{region 'Documentation'}
(*!
<summary>Checks an individually impossible execution budget against actual usable capacity.</summary>
<description>

Real subject boundaries

The real Test Case computes reservations; the real Orchestrator decides and publishes its diagnostic.
A collection double supplies one fixed child view. Only the concurrent Suite allowance is held by
the fixture, without running a Suite. Request-entry observations are inherited from the thin child adapter.
The physical array includes one unused FIFO position, leaving capacity one entry below the minimum.
The buffer is empty at rejection: consumer deletion cannot repair an impossible budget.
Three later helper calls must retain Error without another diagnostic or unexpected dispatch.
Expected diagnostics stay in local capture. The surrounding Assertions use the normal selftest publisher.
The real subject binds only local storage; expected findings remain in that storage.
Checking Assertions retain the outer selftest publisher. Each run reinitializes the subject.
</description>
*)
{endregion}
FUNCTION_BLOCK Test_ImpossibleExecutionBudget EXTENDS TestCaseBase
VAR
    FSubject : EventBuffer;
    FEvents : ARRAY[1..BufferLength] OF ST_Event;
    FFifo : ST_FifoStatus;
    FBufferStatus : ST_EventBufferStatus;
    FPerformed : BOOL;
    FChecked : BOOL;
    FSubjectParent : I_TestSuite;
    FChild : ReservationChildProbe;
    FOrchestrator : OrchestratorProbe;
    FCollection : OrchestrationCollectionDouble;
    FChildren : ARRAY[1..1] OF I_Orchestratable;
    FOwnerReserved : UINT;
    FStep : INT;
    FObservationCalls : UINT;
    FPrecondition : AssertTrue;
    FPreconditionMatches : BOOL;
    FFailureDetection : AssertTrue;
    FFailureDetectionMatches : BOOL;
    FStateAndCounts : AssertTrue;
    FStateAndCountsMatches : BOOL;
    FHeldError : AssertTrue;
    FHeldErrorMatches : BOOL;
    FSingleDiagnostic : AssertTrue;
    FSingleDiagnosticMatches : BOOL;
    FRequestBoundary : AssertTrue;
    FRequestBoundaryMatches : BOOL;
    FAccounting : AssertTrue;
    FAccountingMatches : BOOL;
    FCaptureIntegrity : AssertTrue;
    FCaptureIntegrityMatches : BOOL;
END_VAR
VAR CONSTANT
    ChildExecutionBudget : UINT := 11;
    ConfigureExecution : INT := 4;
    BufferLength : UINT := GVL_Constants.TestSuiteExecutionEventCount + ChildExecutionBudget + Param_EventBuffer.EventBufferExecutionHeadroom;
    ObservationCalls : UINT := 3;
    ExpectedResetRequests : UINT := 1;
    ExpectedStartRequests : UINT := 0;
    Setup : INT := 0;
    PrepareChild : INT := 1;
    TriggerFailure : INT := 2;
    ObserveFailure : INT := 3;
END_VAR

SUPER^();

{region 'Documentation'}
(*!
<summary>Contributes each checking Assertion once.</summary>
*)
{endregion}
METHOD PROTECTED AggregateResults
VAR_INPUT
    Aggregator : I_ResultAggregator; //! Borrowed result sink owned by the outer Test Case; add this test's checking Assertions without resetting or retaining the sink.
END_VAR
Aggregator.AddProvider(Provider := FPrecondition);
Aggregator.AddProvider(Provider := FFailureDetection);
Aggregator.AddProvider(Provider := FStateAndCounts);
Aggregator.AddProvider(Provider := FHeldError);
Aggregator.AddProvider(Provider := FSingleDiagnostic);
Aggregator.AddProvider(Provider := FRequestBoundary);
Aggregator.AddProvider(Provider := FAccounting);
Aggregator.AddProvider(Provider := FCaptureIntegrity);
END_METHOD

{region 'Documentation'}
(*!
<summary>Supplies only the child identity before initialization.</summary>
*)
{endregion}
METHOD PUBLIC BindSubjectParent
VAR_INPUT
    Parent : I_TestSuite; //! Borrowed identity parent retained for isolated subject initialization; keep the Suite alive through subject use.
END_VAR
FSubjectParent := Parent;
END_METHOD

{region 'Documentation'}
(*!
<summary>Calls the real helper and child and retains accounting observations.</summary>
*)
{endregion}
METHOD PRIVATE CallSubject
VAR_INPUT
    Task : E_OrchestratorTask; //! Orchestration task assigned for this controlled subject call.
END_VAR
FOrchestrator(Task := Task);
FAccountingMatches := FAccountingMatches
    AND (FSubject.ReservedEntryCount = FOwnerReserved + FChild.ReservedEntryCount);
FChild();
FCaptureIntegrityMatches := FCaptureIntegrityMatches
    AND NOT FFifo.ConfigError AND NOT FFifo.IndexError
    AND (FBufferStatus.LostEventCount = 0)
    AND NOT FCollection.InvalidAccess AND NOT FCollection.TraceOverflow;
END_METHOD

{region 'Documentation'}
(*!
<summary>Checks the single retained Orchestrator Error and exact dispatch counts.</summary>
*)
{endregion}
METHOD PRIVATE CheckDiagnostic
VAR
    Index : UINT;
    ErrorCount : UINT;
    PayloadMatches : BOOL := TRUE;
END_VAR
FOR Index := 1 TO BufferLength DO
    IF (FEvents[Index].SequenceId > 0) AND (FEvents[Index].Severity = E_EventSeverity.Error) THEN
        ErrorCount := ErrorCount + 1;
        PayloadMatches := PayloadMatches
            AND (FEvents[Index].OwnerScope = E_OwnerScope.Framework)
            AND (FEvents[Index].EventType = E_EventType.Framework)
            AND (FEvents[Index].State = E_State.Error)
            AND (FEvents[Index].Name = CONCAT(Name, '.Orchestrator'))
            AND (FEvents[Index].Message <> '');
    END_IF;
END_FOR;
FSingleDiagnosticMatches := (ErrorCount = 1) AND PayloadMatches;
FRequestBoundaryMatches := FChild.RequestsReserved
    AND (FChild.ResetRequestCount = ExpectedResetRequests)
    AND (FChild.StartRequestCount = ExpectedStartRequests);
END_METHOD

{region 'Documentation'}
(*!
<summary>Requires all checking Assertions to be initialized.</summary>
*)
{endregion}
METHOD PROTECTED CheckInitialization : BOOL //! TRUE when the inherited initialization check and this concrete fixture check both accept the setup.
CheckInitialization := FALSE;
IF NOT SUPER^.CheckInitialization() OR (FSubjectParent = 0) THEN
    RETURN;
END_IF;

CheckInitialization := FPrecondition.IsInitialized
    AND FFailureDetection.IsInitialized
    AND FStateAndCounts.IsInitialized
    AND FHeldError.IsInitialized
    AND FSingleDiagnostic.IsInitialized
    AND FRequestBoundary.IsInitialized
    AND FAccounting.IsInitialized
    AND FCaptureIntegrity.IsInitialized;
END_METHOD

{region 'Documentation'}
(*!
<summary>Initializes the checking Assertions for one test state.</summary>
*)
{endregion}
METHOD PROTECTED Configure
FPreparationStateCount := 0;
FTestStateCount := 1;
FPrecondition.Initialize(Parent := THIS^,
    AssertionName := 'Precondition');
FFailureDetection.Initialize(Parent := THIS^,
    AssertionName := 'FailureDetection');
FStateAndCounts.Initialize(Parent := THIS^,
    AssertionName := 'StateAndCounts');
FHeldError.Initialize(Parent := THIS^,
    AssertionName := 'HeldError');
FSingleDiagnostic.Initialize(Parent := THIS^,
    AssertionName := 'SingleDiagnostic');
FRequestBoundary.Initialize(Parent := THIS^,
    AssertionName := 'RequestBoundary');
FAccounting.Initialize(Parent := THIS^,
    AssertionName := 'Accounting');
FCaptureIntegrity.Initialize(Parent := THIS^,
    AssertionName := 'CaptureIntegrity');
END_METHOD

{region 'Documentation'}
(*!
<summary>Binds a real child and Orchestrator to fixed isolated storage.</summary>
*)
{endregion}
METHOD PRIVATE InitializeArrangement
VAR
    Config : ST_TestCaseConfig;
END_VAR
IF NOT FSubject.Initialize(Buffer := FEvents,
    FifoControl := FFifo,
    Status := FBufferStatus) THEN
    Error(Message := 'Reservation error capture initialization failed.');
    RETURN;
END_IF;
FOwnerReserved := 0;
FChild.BindPublisher(Publisher := FSubject);
FChild.ClearRequestTrace();
FChild.ExecutionSlot := 1;
IF NOT FChild.Initialize(Parent := FSubjectParent,
    TestName := 'ExecutionBudgetChild',
    Config := Config) THEN
    Error(Message := 'Reservation error child initialization failed.');
    RETURN;
END_IF;
FChild();
FChildren[1] := FChild;
IF NOT FCollection.Initialize(Count := 1,
    Children := FChildren) THEN
    Error(Message := 'Reservation error collection initialization failed.');
    RETURN;
END_IF;
FOrchestrator.BindPublisher(Publisher := FSubject);
IF NOT FOrchestrator.Initialize(Collection := FCollection,
    Name := Name) THEN
    Error(Message := 'Reservation error Orchestrator initialization failed.');
    RETURN;
END_IF;
IF NOT FSubject.ReserveSpace(EntryCount := GVL_Constants.TestSuiteResetEventCount,
    HeadroomEntryCount := Param_EventBuffer.EventBufferResetHeadroom,
    OwnerReservedEntryCount := FOwnerReserved) THEN
    Error(Message := 'Reservation error concurrent owner setup failed.');
    RETURN;
END_IF;
FPreconditionMatches := FPreconditionMatches AND FChild.IsInitialized
    AND FFifo.BufferEmpty AND (FSubject.Capacity = BufferLength - 1);
END_METHOD

{region 'Documentation'}
(*!
<summary>Removes setup events and replaces the fixture owner allowance; child configuration remains unchanged.</summary>
*)
{endregion}
METHOD PRIVATE PrepareExecution
VAR
    Watermark : UDINT;
END_VAR
Watermark := FBufferStatus.SequenceId;
FSubject.ProcessDeleteRequest(SequenceId := Watermark);
IF NOT FSubject.FreeReservedSpace(EntryCount := FOwnerReserved,
    OwnerReservedEntryCount := FOwnerReserved) THEN
    Error(Message := 'Could not release Reset fixture allowance.');
    RETURN;
END_IF;
IF NOT FSubject.ReserveSpace(EntryCount := GVL_Constants.TestSuiteExecutionEventCount,
    HeadroomEntryCount := Param_EventBuffer.EventBufferExecutionHeadroom,
    OwnerReservedEntryCount := FOwnerReserved) THEN
    Error(Message := 'Could not reserve execution fixture allowance.');
    RETURN;
END_IF;
FPreconditionMatches := FPreconditionMatches AND FFifo.BufferEmpty
    AND (Watermark = 0) AND (FChild.ReservedEntryCount = 0);
END_METHOD

{region 'Documentation'}
(*!
<summary>Completes abort without asynchronous work.</summary>
*)
{endregion}
METHOD PROTECTED ProcessAbort
VAR_INPUT
    Enable : BOOL; //! Phase permission supplied by the owning Test Case; FALSE does not authorize progression, while observation may continue.
END_VAR
IF Enable THEN
    CompleteAbort();
END_IF;
END_METHOD

{region 'Documentation'}
(*!
<summary>Evaluates captured observations after the scenario has finished.</summary>
*)
{endregion}
METHOD PROTECTED ProcessAssertions
VAR_INPUT
    Enable : BOOL; //! Phase permission supplied by the owning Test Case; FALSE does not authorize progression, while observation may continue.
END_VAR
VAR
    Evaluate : BOOL;
END_VAR
Evaluate := Enable AND FPerformed;
FPrecondition(Enable := Evaluate,
    State := State,
    IN := FPreconditionMatches);
FFailureDetection(Enable := Evaluate,
    State := State,
    IN := FFailureDetectionMatches);
FStateAndCounts(Enable := Evaluate,
    State := State,
    IN := FStateAndCountsMatches);
FHeldError(Enable := Evaluate,
    State := State,
    IN := FHeldErrorMatches);
FSingleDiagnostic(Enable := Evaluate,
    State := State,
    IN := FSingleDiagnosticMatches);
FRequestBoundary(Enable := Evaluate,
    State := State,
    IN := FRequestBoundaryMatches);
FAccounting(Enable := Evaluate,
    State := State,
    IN := FAccountingMatches);
FCaptureIntegrity(Enable := Evaluate,
    State := State,
    IN := FCaptureIntegrityMatches);
IF Evaluate THEN
    FChecked := TRUE;
END_IF;
END_METHOD

{region 'Documentation'}
(*!
<summary>No Preparation phase is needed.</summary>
*)
{endregion}
METHOD PROTECTED ProcessPreparations
VAR_INPUT
    // SA0033: Required override without Preparation work.
    {attribute 'analysis' := '-33'}
    Enable : BOOL; //! Phase permission supplied by the owning Test Case; FALSE does not authorize progression, while observation may continue.
END_VAR
END_METHOD

{region 'Documentation'}
(*!
<summary>Clears scenario evidence; next execution initializes a fresh local arrangement.</summary>
*)
{endregion}
METHOD PROTECTED ProcessReset
FStep := Setup;
FObservationCalls := 0;
FPerformed := FALSE;
FChecked := FALSE;
FPrecondition.Reset();
FPreconditionMatches := TRUE;
FFailureDetection.Reset();
FFailureDetectionMatches := TRUE;
FStateAndCounts.Reset();
FStateAndCountsMatches := TRUE;
FHeldError.Reset();
FHeldErrorMatches := TRUE;
FSingleDiagnostic.Reset();
FSingleDiagnosticMatches := TRUE;
FRequestBoundary.Reset();
FRequestBoundaryMatches := TRUE;
FAccounting.Reset();
FAccountingMatches := TRUE;
FCaptureIntegrity.Reset();
FCaptureIntegrityMatches := TRUE;
FSingleDiagnosticMatches := FALSE;
CompleteReset();
END_METHOD

{region 'Documentation'}
(*!
<summary>Advances one scenario phase before checking final captured observations.</summary>
*)
{endregion}
METHOD PROTECTED ProcessTests
VAR_INPUT
    Enable : BOOL; //! Phase permission supplied by the owning Test Case; FALSE does not authorize progression, while observation may continue.
END_VAR
IF NOT Enable THEN
    RETURN;
END_IF;
IF FChecked THEN
    CompleteTests();
    RETURN;
END_IF;
IF NOT FPerformed THEN
    RunScenario();
END_IF;
END_METHOD

{region 'Documentation'}
(*!
<summary>Runs one bounded scenario phase per active outer call.</summary>
*)
{endregion}
METHOD PRIVATE RunScenario
CASE FStep OF
    Setup:
        InitializeArrangement();
        FStep := PrepareChild;

    PrepareChild:
        CallSubject(Task := E_OrchestratorTask.Reset);
        IF FOrchestrator.Result = E_Result.Error THEN
            Error(Message := 'Reservation error scenario could not reset its child.');
            RETURN;
        END_IF;
        IF FOrchestrator.IsResetFinished THEN
            FPreconditionMatches := FPreconditionMatches AND FChild.IsIdle AND FChild.IsReady;
            FStep := ConfigureExecution;
        END_IF;

    ConfigureExecution:
        CallSubject(Task := E_OrchestratorTask.Idle);
        PrepareExecution();
        FStep := TriggerFailure;

    TriggerFailure:
        TriggerSubjectFailure();
        FStep := ObserveFailure;

    ObserveFailure:
        CallSubject(Task := E_OrchestratorTask.Execution);
        FFailureDetectionMatches := FFailureDetectionMatches
            AND (FOrchestrator.Result = E_Result.Error);
        FHeldErrorMatches := FHeldErrorMatches
            AND (FOrchestrator.Result = E_Result.Error)
            AND NOT FOrchestrator.IsExecutionFinished;
        FObservationCalls := FObservationCalls + 1;
        IF FObservationCalls = ObservationCalls THEN
            CheckDiagnostic();
            FAccountingMatches := FAccountingMatches
                AND (FChild.ReservedEntryCount = 0);
            IF NOT FSubject.FreeReservedSpace(EntryCount := FOwnerReserved,
                OwnerReservedEntryCount := FOwnerReserved) THEN
                Error(Message := 'Reservation error fixture cleanup failed.');
                RETURN;
            END_IF;
            FAccountingMatches := FAccountingMatches AND (FSubject.ReservedEntryCount = 0);
            FPerformed := TRUE;
        END_IF;
ELSE
    Error(Message := 'Unknown reservation error test step.');
END_CASE;
END_METHOD

{region 'Documentation'}
(*!
<summary>Classifies the impossible budget on an empty buffer, then exercises real Orchestrator handling.</summary>
*)
{endregion}
METHOD PRIVATE TriggerSubjectFailure
VAR
    ReservationResult : E_EventReservationResult;
    PreviousSequence : UDINT;
    PreviousState : E_State;
END_VAR
PreviousSequence := FBufferStatus.SequenceId;
PreviousState := FChild.State;
ReservationResult := FChild.ReserveExecutionEvents();
FFailureDetectionMatches := ReservationResult = E_EventReservationResult.Error;
FStateAndCountsMatches := (FChild.State = PreviousState)
    AND (FChild.ReservedEntryCount = 0)
    AND (FSubject.ReservedEntryCount = FOwnerReserved)
    AND (FBufferStatus.SequenceId = PreviousSequence)
    AND FFifo.BufferEmpty;
CallSubject(Task := E_OrchestratorTask.Execution);
FFailureDetectionMatches := FFailureDetectionMatches
    AND (FOrchestrator.Result = E_Result.Error);
END_METHOD

END_FUNCTION_BLOCK

(* stored: Version 1.1.0.1
   POU Test_ImpossibleExecutionBudget: Id {daf0992d-343d-4dfb-a1fa-6c5108466c62}, SpecialFunc None
   Folder Internal: Id {037d414a-5282-4206-910a-1821eccd8192}
   Method AggregateResults: Id {a963fca6-db4f-4bd3-8f92-6108d1e4a5a9}
   Method BindSubjectParent: Id {d0604b6d-c7cf-4fe0-8673-016ebbc2f184}
   Method CallSubject: Id {a8baa7d7-e6a2-43f1-959d-8261a6e22e88}
   Method CheckDiagnostic: Id {95faac6f-201a-437a-81a4-b41aef5b866e}
   Method CheckInitialization: Id {d9267834-bdb1-4ae3-88e3-df8d39e290c2}
   Method Configure: Id {a713066b-5016-4aba-9c4d-ddc933b38826}
   Method InitializeArrangement: Id {a8f9048e-cf62-4fbd-85b6-75d8dff7b296}
   Method PrepareExecution: Id {84d9f129-a27d-499e-95b5-436c955c1824}
   Method ProcessAbort: Id {8c7c72e9-b7fe-418a-a3e5-5a4054301f93}
   Method ProcessAssertions: Id {2cc98cf9-e6e7-4029-8024-e878c6d52e7f}
   Method ProcessPreparations: Id {0ce8be0f-330e-4a39-a5bd-592f442c019b}
   Method ProcessReset: Id {a8386674-13a1-49fe-bbbc-fd6137da1353}
   Method ProcessTests: Id {85384ad7-02f3-4410-800e-a66ae870fe37}
   Method RunScenario: Id {6a1be4a9-c370-4540-b0b7-534c26661b95}
   Method TriggerSubjectFailure: Id {e9991f6c-1515-49b2-8125-c1b45ef5e66f} *)
